FUNCTION_BLOCK FB_CoverOpeningState EXTENDS FB_CoverState
VAR
	nStage			: UINT:= 0;
	tonDelta		: TON;		// PT is taken from pCover^.Delta at the start of each cycle (#76)
	tonFullCycle	: TON;		// PT is taken from pCover^.TimeToCycle at the start of each cycle (#76)
END_VAR

METHOD CloseCommand : BOOL
nStage := 0;
tonDelta(IN:=FALSE);
tonFullCycle(IN:=FALSE);
pCover^.SetState(pCover^.fbCoverClosingState);
END_METHOD

METHOD RunState : BOOL
tonDelta();
tonFullCycle();
CASE nStage OF
	0:
		// #76: the cycle times were only read once, by the declaration initialisers, so the inputs of FB_CoverControl
		// never reached the timers. Take them at the start of each cycle (not every scan: a change mid-cycle must not
		// end it early).
		tonDelta.PT := pCover^.Delta;
		IF pCover^.TimeToCycle > T#0S THEN
			tonFullCycle.PT := pCover^.TimeToCycle;
		ELSE
			tonFullCycle.PT := T#15S;	// 0 would declare the end position after one scan
		END_IF
		pCover^._CoverState := E_MirrorCoverState.opening;
		tonDelta.IN:=TRUE;
		nStage := 1;
	1:
		// Open Motor 1
		pCover^._Motor1RelaisA := TRUE;
		pCover^._Motor1RelaisB := FALSE;
		// Stop Motor 2
		pCover^._Motor2RelaisA := FALSE;
		pCover^._Motor2RelaisB := FALSE;
		nStage := 2;
	2:
		IF tonDelta.Q THEN
			tonDelta.IN:=FALSE;
			nStage:=3;
		END_IF 
	3:
		// Open Motor 2
		pCover^._Motor2RelaisA := TRUE;
		pCover^._Motor2RelaisB := FALSE;
		tonFullCycle.IN:=TRUE;
		nStage := 4;
	4:
		IF tonFullCycle.Q THEN
			tonFullCycle.IN:=FALSE;
			THIS^.SuccessfulFinished();
		END_IF 
END_CASE
END_METHOD

METHOD StopCommand : BOOL
nStage := 0;
tonDelta(IN:=FALSE);
tonFullCycle(IN:=FALSE);
pCover^.SetState(pCover^.fbCoverStoppingState);
END_METHOD

METHOD SuccessfulFinished : BOOL
nStage := 0;
tonDelta(IN:=FALSE);
tonFullCycle(IN:=FALSE);
// #71: release the relays at the end position (limit switches cut the motors, the covers are self-locking)
pCover^._Motor1RelaisA := FALSE;
pCover^._Motor1RelaisB := FALSE;
pCover^._Motor2RelaisA := FALSE;
pCover^._Motor2RelaisB := FALSE;
pCover^._CoverState := E_MirrorCoverState.open;
pCover^.SetState(pCover^.fbCoverIdleState);
END_METHOD

END_FUNCTION_BLOCK

(* stored: Version 1.1.0.1, ProductVersion 3.1.4024.15
   POU FB_CoverOpeningState: Id {f67eb63e-4b73-4ad7-b7b5-3044d6304760}, SpecialFunc None
   Method CloseCommand: Id {099c7f81-ac72-43ae-9efb-0a90bfcce006}
   Method RunState: Id {89fa8360-8bdf-4734-ab38-105f69dc24d7}
   Method StopCommand: Id {30bb32b5-d910-4771-948e-56435f53e601}
   Method SuccessfulFinished: Id {cfd5f6a0-880a-440e-9a62-ea7a6ddf139e} *)
